FUNCTION_BLOCK Controller (* Extracted Composite Function Block Type *)
  (* Version 3/26/2020, prana *)
  PACKAGE Main;
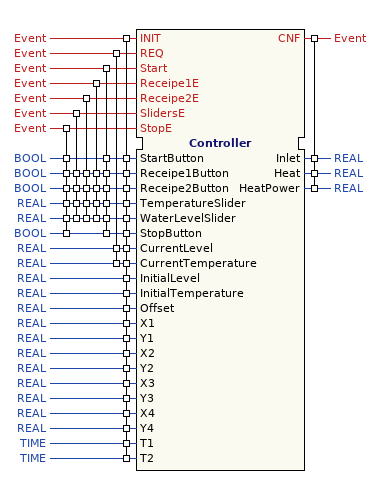
  EVENT_INPUT
    INIT WITH StartButton, Receipe1Button, Receipe2Button, TemperatureSlider, WaterLevelSlider, StopButton, CurrentLevel, CurrentTemperature, InitialLevel, InitialTemperature, Offset, Y2, X3, Y3, X4, Y4, T1, T2, X1, Y1, X2;
    REQ WITH CurrentTemperature, CurrentLevel; (* Normal Execution Request *)
    Start WITH StartButton, Receipe1Button, Receipe2Button, TemperatureSlider, WaterLevelSlider, StopButton;
    Receipe1E WITH Receipe1Button, Receipe2Button, TemperatureSlider, WaterLevelSlider; (* Initialization Request *)
    Receipe2E WITH Receipe1Button, Receipe2Button, TemperatureSlider, WaterLevelSlider; (* Normal Execution Request *)
    SlidersE WITH Receipe1Button, Receipe2Button, TemperatureSlider, WaterLevelSlider;
    StopE WITH StartButton, Receipe1Button, Receipe2Button, TemperatureSlider, WaterLevelSlider, StopButton;
  END_EVENT
  EVENT_OUTPUT
    CNF WITH Inlet, Heat, HeatPower; (* Execution Confirmation *)
  END_EVENT
  VAR_INPUT
    StartButton : BOOL;
    Receipe1Button : BOOL; (* Input event qualifier *)
    Receipe2Button : BOOL;
    TemperatureSlider : REAL;
    WaterLevelSlider : REAL;
    StopButton : BOOL;
    CurrentLevel : REAL; (* Input event qualifier *)
    CurrentTemperature : REAL; (* Input event qualifier *)
    InitialLevel : REAL;
    InitialTemperature : REAL;
    Offset : REAL;
    X1 : REAL;
    Y1 : REAL;
    X2 : REAL;
    Y2 : REAL;
    X3 : REAL;
    Y3 : REAL;
    X4 : REAL;
    Y4 : REAL;
    T1 : TIME;
    T2 : TIME;
  END_VAR
  VAR_OUTPUT
    Inlet : REAL; (* Output event qualifier *)
    Heat : REAL;
    HeatPower : REAL;
  END_VAR
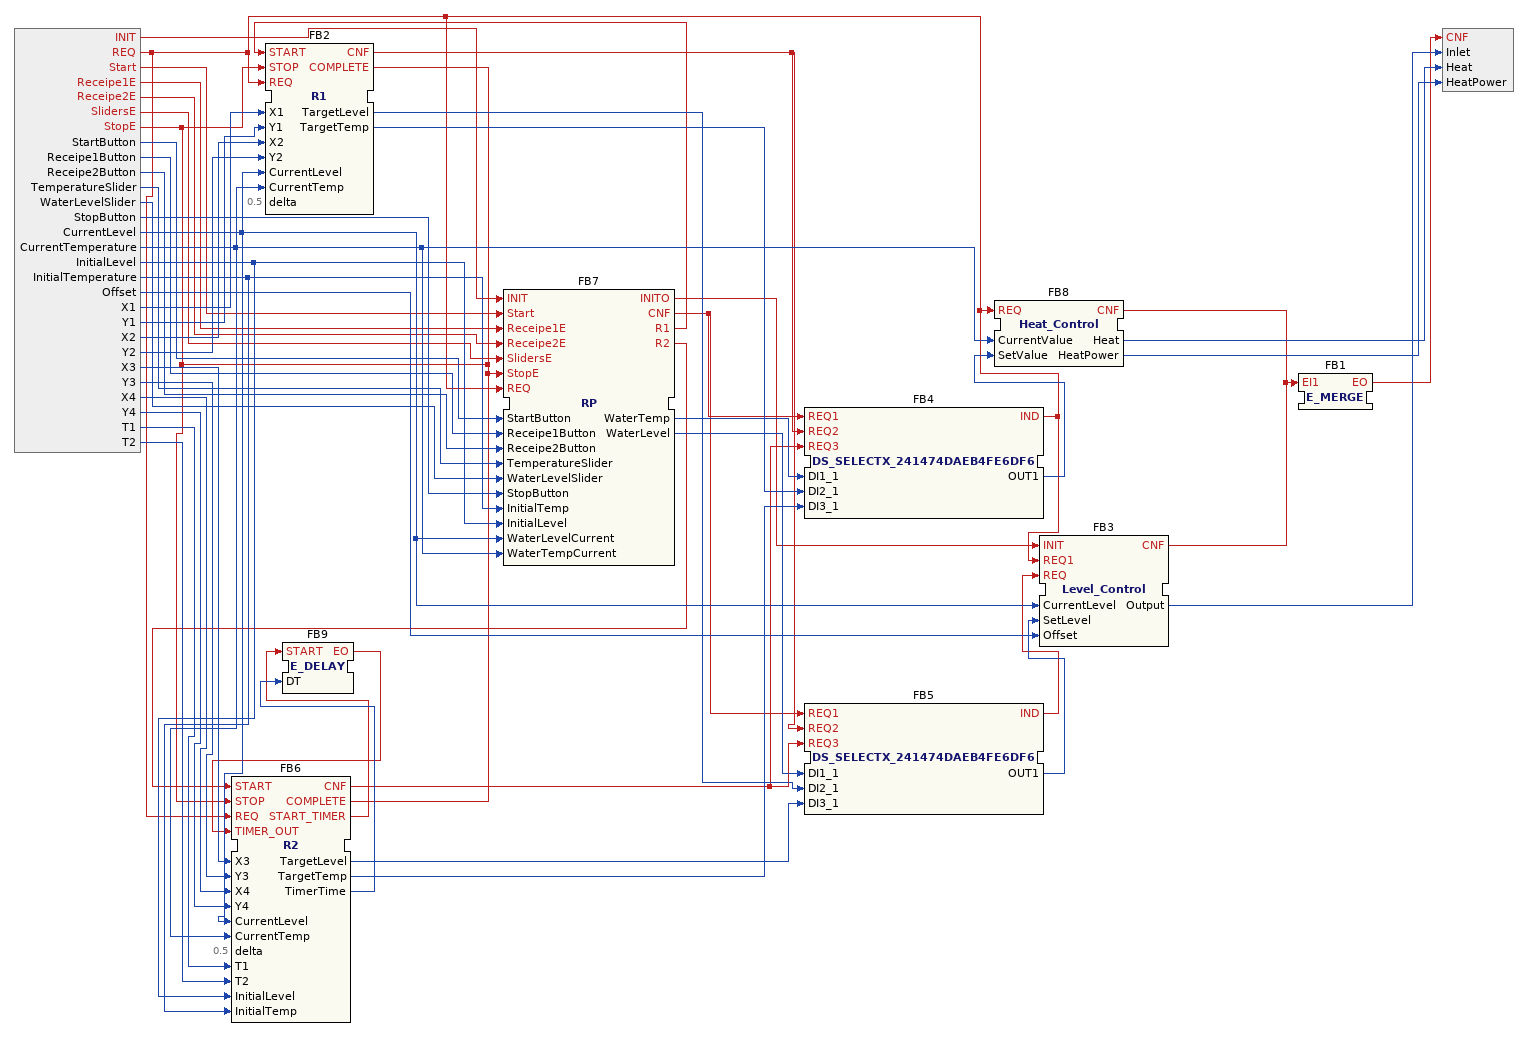
  FBS
    FB7 : RP;
    FB8 : Heat_Control;
    FB3 : Level_Control;
    FB1 : E_MERGE;
    FB2 : R1(delta := 0.5);
    FB4 : DS_SELECTX_241474DAEB4FE6DF6; {SET_ATTRIBUTE(Configuration.GenericFBType.InterfaceParams, Runtime.Standard#CNTX:=3;CNTY:=1;DI${CNTX,_,CNTY$}:REAL)}
    FB5 : DS_SELECTX_241474DAEB4FE6DF6; {SET_ATTRIBUTE(Configuration.GenericFBType.InterfaceParams, Runtime.Standard#CNTX:=3;CNTY:=1;DI${CNTX,_,CNTY$}:REAL)}
    FB6 : R2(delta := 0.5);
    FB9 : E_DELAY;
  END_FBS
  EVENT_CONNECTIONS
    FB7.INITO TO FB3.INIT;
    Start TO FB7.Start;
    Receipe1E TO FB7.Receipe1E;
    Receipe2E TO FB7.Receipe2E;
    SlidersE TO FB7.SlidersE;
    StopE TO FB7.StopE;
    REQ TO FB8.REQ;
    REQ TO FB3.REQ1;
    REQ TO FB7.REQ;
    FB8.CNF TO FB1.EI1;
    FB3.CNF TO FB1.EI1;
    FB1.EO TO CNF;
    INIT TO FB7.INIT;
    FB7.R1 TO FB2.START;
    StopE TO FB2.STOP;
    REQ TO FB2.REQ;
    FB2.COMPLETE TO FB7.StopE;
    FB7.R2 TO FB6.START;
    StopE TO FB6.STOP;
    FB6.COMPLETE TO FB7.StopE;
    FB7.CNF TO FB5.REQ1;
    FB2.CNF TO FB5.REQ2;
    FB5.IND TO FB3.REQ;
    FB6.CNF TO FB5.REQ3;
    FB7.CNF TO FB4.REQ1;
    FB2.CNF TO FB4.REQ2;
    FB4.IND TO FB8.REQ;
    FB6.CNF TO FB4.REQ3;
    FB6.START_TIMER TO FB9.START;
    FB9.EO TO FB6.TIMER_OUT;
    REQ TO FB6.REQ;
  END_CONNECTIONS
  DATA_CONNECTIONS
    StartButton TO FB7.StartButton;
    Receipe1Button TO FB7.Receipe1Button;
    Receipe2Button TO FB7.Receipe2Button;
    TemperatureSlider TO FB7.TemperatureSlider;
    WaterLevelSlider TO FB7.WaterLevelSlider;
    StopButton TO FB7.StopButton;
    CurrentTemperature TO FB8.CurrentValue;
    FB8.Heat TO Heat;
    CurrentLevel TO FB3.CurrentLevel;
    FB3.Output TO Inlet;
    CurrentTemperature TO FB7.WaterTempCurrent;
    CurrentLevel TO FB7.WaterLevelCurrent;
    InitialLevel TO FB7.InitialLevel;
    InitialTemperature TO FB7.InitialTemp;
    FB8.HeatPower TO HeatPower;
    Offset TO FB3.Offset;
    CurrentLevel TO FB2.CurrentLevel;
    CurrentTemperature TO FB2.CurrentTemp;
    X1 TO FB2.X1;
    Y1 TO FB2.Y1;
    X2 TO FB2.X2;
    Y2 TO FB2.Y2;
    InitialTemperature TO FB6.InitialTemp;
    InitialLevel TO FB6.InitialLevel;
    X3 TO FB6.X3;
    Y3 TO FB6.Y3;
    X4 TO FB6.X4;
    Y4 TO FB6.Y4;
    T1 TO FB6.T1;
    T2 TO FB6.T2;
    CurrentLevel TO FB6.CurrentLevel;
    CurrentTemperature TO FB6.CurrentTemp;
    FB7.WaterLevel TO FB5.DI1_1;
    FB2.TargetLevel TO FB5.DI2_1;
    FB5.OUT1 TO FB3.SetLevel;
    FB6.TargetLevel TO FB5.DI3_1;
    FB7.WaterTemp TO FB4.DI1_1;
    FB2.TargetTemp TO FB4.DI2_1;
    FB4.OUT1 TO FB8.SetValue;
    FB6.TargetTemp TO FB4.DI3_1;
    FB6.TimerTime TO FB9.DT;
  END_CONNECTIONS
END_FUNCTION_BLOCK
